// // MIGRATION DRAFT: not included in PLC compilation.
// // Reference: Reference_Project/VTD_HMI_FB.scl, object VTD_HMI_FB.
// // Types, globals, calls, units and behavior require manual reconciliation.
// // See docs/TIA_Missing_Blocks.md before importing as PLC code.
FUNCTION_BLOCK VTD_HMI_FB
// 
//    VAR
//       T_Charge   : TON;
//    END_VAR

// // MIGRATION DRAFT: not included in PLC compilation.
// // Reference: Reference_Project/VTD_HMI_FB.scl, object VTD_HMI_FB.
// // Types, globals, calls, units and behavior require manual reconciliation.
// // See docs/TIA_Missing_Blocks.md before importing as PLC code.
// IF VTDtem_Selected_HMI <> VTD_ID_HMI_OLD THEN
// 	    Screen_DB.Charge_VTD_Commands := TRUE;
// 	    VTD_ID_HMI_OLD := VTDtem_Selected_HMI;
// 	END_IF;
// 
// 
// 	IF Screen_DB.Charge_VTD_Commands THEN
// 	    CASE VTDtem_Selected_HMI OF
// 	        1:
// 	            VTD_Mode_Change_HMI := Control.VTD.Mode;
// 	            VTD_Enable_HMI := Control.VTD.Instruction.Enable;
// 	            LE_Bypass := LE_Bypass_1_;
// 	            VTD_Stop_HMI := Control.VTD.Instruction.Stop;
// 	        2:
// 	            VTD_Mode_Change_HMI := Control.VTD[2].Mode;
// 	            VTD_Enable_HMI := Control.VTD[2].Instruction.Enable;
// 	            LE_Bypass := LE_Bypass_2_;
// 	            VTD_Stop_HMI := Control.VTD[2].Instruction.Stop;
// 	        3:
// 	            VTD_Mode_Change_HMI := Control.VTD[3].Mode;
// 	            VTD_Enable_HMI := Control.VTD[3].Instruction.Enable;
// 	            LE_Bypass := LE_Bypass_3_;
// 	            VTD_Stop_HMI := Control.VTD[3].Instruction.Stop;
// 	        4:
// 	            VTD_Mode_Change_HMI := Control.VTD[4].Mode;
// 	            VTD_Enable_HMI := Control.VTD[4].Instruction.Enable;
// 	            LE_Bypass := LE_Bypass_4_;
// 	            VTD_Stop_HMI := Control.VTD[4].Instruction.Stop;
// 	        5:
// 	            VTD_Mode_Change_HMI := Control.VTD[5].Mode;
// 	            VTD_Enable_HMI := Control.VTD[5].Instruction.Enable;
// 	            LE_Bypass := LE_Bypass_5_;
// 	            VTD_Stop_HMI := Control.VTD[5].Instruction.Stop;
// 	    END_CASE;
// 
// 	    T_Charge.TON(IN := TRUE,
// 	                  PT := T#500mS);
// 	    IF T_Charge.Q THEN
// 	        T_Charge.TON(IN := FALSE,
// 	                      PT := T#0mS);
// 	        Screen_DB.Charge_VTD_Commands := 0;
// 	    END_IF;
// 
// 
// 	ELSIF HMI_DB.ScreenNo_Main = 1 AND NOT Screen_DB.Charge_VTD_Commands THEN
// 	    CASE VTDtem_Selected_HMI OF
// 	        1:
// 	            Feed_VTD_HMI_FC(Sys_No := 1,
// 	                              Rem_Loc_Keys:= HMI_DB.Rem_Loc_Keys[1].Level,
// 	                              Safety_OK := Remote_Panel_DB_1.Safety_OK,
// 	                              BCD_Test_Ok_HMI := SICK_Lector_DB_1.Test_OK,
// 	                              BCD_Error_HMI := SICK_Lector_DB_1.Error,
// 	                              BCD_RdDone := SICK_Lector_DB_1.RdDone,
// 	                              BCD_ReqDone := SICK_Lector_DB_1.ReqDone,
// 	                              BCD_ReqBusy := SICK_Lector_DB_1.ReqBusy,
// 	                              Start_InBarcodeStation := Start_InBarcodeStation_HMI,
// 	                              Sick_Lector_Reseult := SICK_Lector_DB_1.Barcode_Result,
// 	                              Level_Below_Extractor := VTD_FB_DB_1.LevelBelowExtractor,
// 	                              Speed_mm_s := VTD_FB_DB_1.VTDSpeed_mm_s,
// 	                              LE_Bypass := LE_Bypass_1_,
// 	                              BCD_Start_Comm_Test_HMI := BCD_Test_Comm_HMI_1_,
// 	                              BCD_Enable_Trigger_HMI := BCD_Enable_Trigger_HMI_1_,
// 	                              BCD_Disable_Trigger_HMI := BCD_Disable_Trigger_HMI_1_,
// 	                              BCD_Execute_Function := SICK_Lector_Control_1.Enable_Req,
// 	                              System_Busy => System_1_Busy);
// 
// 	        2:
// 	            Feed_VTD_HMI_FC(Sys_No := 2,
// 	                              Rem_Loc_Keys:=HMI_DB.Rem_Loc_Keys[2].Level,
// 	                              Safety_OK := Remote_Panel_DB_2.Safety_OK,
// 	                              BCD_Test_Ok_HMI := SICK_Lector_DB_2.Test_OK,
// 	                              BCD_Error_HMI := SICK_Lector_DB_2.Error,
// 	                              BCD_RdDone := SICK_Lector_DB_2.RdDone,
// 	                              BCD_ReqDone := SICK_Lector_DB_2.ReqDone,
// 	                              BCD_ReqBusy := SICK_Lector_DB_2.ReqBusy,
// 	                              Start_InBarcodeStation := Start_InBarcodeStation_HMI,
// 	                              Sick_Lector_Reseult := SICK_Lector_DB_2.Barcode_Result,
// 	                              Level_Below_Extractor := VTD_FB_DB_2.LevelBelowExtractor,
// 	                              Speed_mm_s := VTD_FB_DB_2.VTDSpeed_mm_s,
// 	                              LE_Bypass := LE_Bypass_2_,
// 	                              BCD_Start_Comm_Test_HMI := BCD_Test_Comm_HMI_2_,
// 	                              BCD_Enable_Trigger_HMI := BCD_Enable_Trigger_HMI_2_,
// 	                              BCD_Disable_Trigger_HMI := BCD_Disable_Trigger_HMI_2_,
// 	                              BCD_Execute_Function := SICK_Lector_Control_2.Enable_Req,
// 	                              System_Busy => System_2_Busy);
// 	        3:
// 	            Feed_VTD_HMI_FC(Sys_No := 3,
// 	                              Rem_Loc_Keys:=HMI_DB.Rem_Loc_Keys[3].Level,
// 	                              Safety_OK := Remote_Panel_DB_3.Safety_OK,
// 	                              BCD_Test_Ok_HMI := SICK_Lector_DB_3.Test_OK,
// 	                              BCD_Error_HMI := SICK_Lector_DB_3.Error,
// 	                              BCD_RdDone := SICK_Lector_DB_3.RdDone,
// 	                              BCD_ReqDone := SICK_Lector_DB_3.ReqDone,
// 	                              BCD_ReqBusy := SICK_Lector_DB_3.ReqBusy,
// 	                              Start_InBarcodeStation := Start_InBarcodeStation_HMI,
// 	                              Sick_Lector_Reseult := SICK_Lector_DB_3.Barcode_Result,
// 	                              Level_Below_Extractor := VTD_FB_DB_3.LevelBelowExtractor,
// 	                              Speed_mm_s := VTD_FB_DB_3.VTDSpeed_mm_s,
// 	                              LE_Bypass := LE_Bypass_3_,
// 	                              BCD_Start_Comm_Test_HMI := BCD_Test_Comm_HMI_3_,
// 	                              BCD_Enable_Trigger_HMI := BCD_Enable_Trigger_HMI_3_,
// 	                              BCD_Disable_Trigger_HMI := BCD_Disable_Trigger_HMI_3_,
// 	                              BCD_Execute_Function := SICK_Lector_Control_3.Enable_Req,
// 	                              System_Busy => System_3_Busy);
// 	        4:
// 	            Feed_VTD_HMI_FC(Sys_No := 4,
// 	                              Rem_Loc_Keys:=HMI_DB.Rem_Loc_Keys[4].Level,
// 	                              Safety_OK := Remote_Panel_DB_4.Safety_OK,
// 	                              BCD_Test_Ok_HMI := SICK_Lector_DB_4.Test_OK,
// 	                              BCD_Error_HMI := SICK_Lector_DB_4.Error,
// 	                              BCD_RdDone := SICK_Lector_DB_4.RdDone,
// 	                              BCD_ReqDone := SICK_Lector_DB_4.ReqDone,
// 	                              BCD_ReqBusy := SICK_Lector_DB_4.ReqBusy,
// 	                              Start_InBarcodeStation := Start_InBarcodeStation_HMI,
// 	                              Sick_Lector_Reseult := SICK_Lector_DB_4.Barcode_Result,
// 	                              Level_Below_Extractor := VTD_FB_DB_4.LevelBelowExtractor,
// 	                              Speed_mm_s := VTD_FB_DB_4.VTDSpeed_mm_s,
// 	                              LE_Bypass := LE_Bypass_4_,
// 	                              BCD_Start_Comm_Test_HMI := BCD_Test_Comm_HMI_4_,
// 	                              BCD_Enable_Trigger_HMI := BCD_Enable_Trigger_HMI_4_,
// 	                              BCD_Disable_Trigger_HMI := BCD_Disable_Trigger_HMI_4_,
// 	                              BCD_Execute_Function := SICK_Lector_Control_4.Enable_Req,
// 	                              System_Busy => System_4_Busy);
// 	        5:
// 	            Feed_VTD_HMI_FC(Sys_No := 5,
// 	                              Rem_Loc_Keys:=HMI_DB.Rem_Loc_Keys[5].Level,
// 	                              Safety_OK := Remote_Panel_DB_5.Safety_OK,
// 	                              BCD_Test_Ok_HMI := SICK_Lector_DB_5.Test_OK,
// 	                              BCD_Error_HMI := SICK_Lector_DB_5.Error,
// 	                              BCD_RdDone := SICK_Lector_DB_5.RdDone,
// 	                              BCD_ReqDone := SICK_Lector_DB_5.ReqDone,
// 	                              BCD_ReqBusy := SICK_Lector_DB_5.ReqBusy,
// 	                              Start_InBarcodeStation := Start_InBarcodeStation_HMI,
// 	                              Sick_Lector_Reseult := SICK_Lector_DB_5.Barcode_Result,
// 	                              Level_Below_Extractor := VTD_FB_DB_5.LevelBelowExtractor,
// 	                              Speed_mm_s := VTD_FB_DB_5.VTDSpeed_mm_s,
// 	                              LE_Bypass := LE_Bypass_5_,
// 	                              BCD_Start_Comm_Test_HMI := BCD_Test_Comm_HMI_5_,
// 	                              BCD_Enable_Trigger_HMI := BCD_Enable_Trigger_HMI_5_,
// 	                              BCD_Disable_Trigger_HMI := BCD_Disable_Trigger_HMI_5_,
// 	                              BCD_Execute_Function := SICK_Lector_Control_5.Enable_Req,
// 	                              System_Busy => System_5_Busy);
// 	    END_CASE;
// 	END_IF;

END_FUNCTION_BLOCK

(* stored: Version 1.1.0.1
   POU VTD_HMI_FB: Id {854ba2e1-d64b-5b2c-b84f-5cc925c23140}, SpecialFunc None *)
